KUKA KRL program: WeldingAddin.src

&ACCESS RVP
&REL 1
&PARAM TEMPLATE = C:\KRC\Roboter\Template\vorgabe
&PARAM EDITMASK = *
DEF WeldingAddin ( )

;FOLD INI
  ;FOLD BASISTECH INI
    GLOBAL INTERRUPT DECL 3 WHEN $STOPMESS==TRUE DO IR_STOPM ( )
    INTERRUPT ON 3
    BAS (#INITMOV,0 )
  ;ENDFOLD (BASISTECH INI)




;FOLD ARCTECH_ANALOG INI
IF A10_OPTION==#ACTIVE THEN
INTERRUPT DECL A_Arc_Control_Intr WHEN $CYCFLAG[A_CycFlagIndex1]==FALSE DO A10 (#APPL_ERROR)
INTERRUPT DECL A_Arc_Swi_Intr WHEN A_ARC_SWI==#ACTIVE DO A10 (#ARC_SEAM)
INTERRUPT DECL A_Arc_HPU_Intr WHEN A_FLY_ARC==TRUE DO A10 (#HPU_ARC)
INTERRUPT  ON A_Arc_HPU_Intr
A10_INI ( )
ENDIF
;ENDFOLD (ARCTECH_ANALOG INI)
  ;FOLD USER INI
        ;FOLD SAFETY HOLDER INI
GLOBAL INTERRUPT DECL 5 WHEN $IN[5]==FALSE DO SAFETY_HOLDER()
INTERRUPT ON 5

;ENDFOLD (SAFETY HOLDER INI)
    ;Make your modifications here

  ;ENDFOLD (USER INI)
;ENDFOLD (INI)
;FOLD PTP HOME Vel=20 % DEFAULT;%{PE}%R 5.6.13,%MKUKATPBASIS,%CMOVE,%VPTP,%P 1:PTP, 2:HOME, 3:, 5:20, 7:DEFAULT
$BWDSTART=FALSE
PDAT_ACT=PDEFAULT
FDAT_ACT=FHOME
BAS(#PTP_PARAMS,20)
$H_POS=XHOME
PTP XHOME
;ENDFOLD



; Program generated by RoboDK v5.7.3 for RoboDK Industrial on 02/07/2024 19:37:37
; Using nominal kinematics.
; Message if failed, eg: Install the Welding Addin
; Message if failed, eg: Install the Welding Addin
BASE_DATA[0] = {FRAME: X 0.000,Y 0.000,Z 0.000,A 0.000,B 0.000,C 0.000}
TOOL_DATA[1] = {FRAME: X 129.073,Y 0.000,Z 85.477,A 0.000,B 22.849,C 0.000}
;FOLD PTP P1 Vel=100.000 % PDAT1 Tool[1] Base[0];%{PE}%R 5.5.31,%MKUKATPBASIS,%CMOVE,%VPTP,%P 1:PTP, 2:P1, 3:, 5:100.000, 7:PDAT1
$BWDSTART=FALSE
PDAT_ACT=PPDAT1
FDAT_ACT=FP1
BAS(#PTP_PARAMS,100)
PTP XP1 C_PTP
;ENDFOLD

; Message if failed, eg: Install the Welding Addin
;FOLD PTP P2 Vel=100.000 % PDAT2 Tool[1] Base[0];%{PE}%R 5.5.31,%MKUKATPBASIS,%CMOVE,%VPTP,%P 1:PTP, 2:P2, 3:, 5:100.000, 7:PDAT2
$BWDSTART=FALSE
PDAT_ACT=PPDAT2
FDAT_ACT=FP2
BAS(#PTP_PARAMS,100)
PTP XP2 C_PTP
;ENDFOLD

;FOLD LIN P3 Vel=1.000 m/s CPDAT3 Tool[1] Base[0];%{PE}%R 5.5.0,%MKUKATPA20,%CARC_SWI,%VLIN,%P 1:LIN, 2:P3, 3:, 5:1.000, 7:CPDAT3
$BWDSTART=FALSE
LDAT_ACT=LCPDAT3
FDAT_ACT=FP3
BAS(#CP_PARAMS,1.000)
LIN XP3 C_DIS
;ENDFOLD

; Message if failed, eg: Install the Welding Addin
;FOLD PTP P4 Vel=100.000 % PDAT4 Tool[1] Base[0];%{PE}%R 5.5.31,%MKUKATPBASIS,%CMOVE,%VPTP,%P 1:PTP, 2:P4, 3:, 5:100.000, 7:PDAT4
$BWDSTART=FALSE
PDAT_ACT=PPDAT4
FDAT_ACT=FP4
BAS(#PTP_PARAMS,100)
PTP XP4 C_PTP
;ENDFOLD

; Previous line is a comment!
; Message if failed, eg: Install the Welding Addin
; Message if failed, eg: Install the Welding Addin
;FOLD PTP P5 Vel=100.000 % PDAT5 Tool[1] Base[0];%{PE}%R 5.5.31,%MKUKATPBASIS,%CMOVE,%VPTP,%P 1:PTP, 2:P5, 3:, 5:100.000, 7:PDAT5
$BWDSTART=FALSE
PDAT_ACT=PPDAT5
FDAT_ACT=FP5
BAS(#PTP_PARAMS,100)
PTP XP5 C_PTP
;ENDFOLD

; Previous line is a comment!
; Message if failed, eg: Install the Welding Addin
;FOLD PTP P6 Vel=100.000 % PDAT6 Tool[1] Base[0];%{PE}%R 5.5.31,%MKUKATPBASIS,%CMOVE,%VPTP,%P 1:PTP, 2:P6, 3:, 5:100.000, 7:PDAT6
$BWDSTART=FALSE
PDAT_ACT=PPDAT6
FDAT_ACT=FP6
BAS(#PTP_PARAMS,100)
PTP XP6 C_PTP
;ENDFOLD

;FOLD LIN P7 Vel=1.000 m/s CPDAT7 Tool[1] Base[0];%{PE}%R 5.5.0,%MKUKATPA20,%CARC_SWI,%VLIN,%P 1:LIN, 2:P7, 3:, 5:1.000, 7:CPDAT7
$BWDSTART=FALSE
LDAT_ACT=LCPDAT7
FDAT_ACT=FP7
BAS(#CP_PARAMS,1.000)
LIN XP7 C_DIS
;ENDFOLD

; Previous line is a comment!
; Message if failed, eg: Install the Welding Addin
; Previous line is a comment!
;FOLD PTP P8 Vel=100.000 % PDAT8 Tool[1] Base[0];%{PE}%R 5.5.31,%MKUKATPBASIS,%CMOVE,%VPTP,%P 1:PTP, 2:P8, 3:, 5:100.000, 7:PDAT8
$BWDSTART=FALSE
PDAT_ACT=PPDAT8
FDAT_ACT=FP8
BAS(#PTP_PARAMS,100)
PTP XP8 C_PTP
;ENDFOLD

END
